FUNCTION F_RealToBitDword_1 : DWORD
VAR_INPUT
	rIn : REAL;
END_VAR
VAR
	pt : POINTER TO DWORD;
END_VAR

pt := ADR(rIn);
F_RealToBitDword := pt^;

END_FUNCTION

(* stored: Version 1.1.0.1, ProductVersion 3.1.4024.15
   POU F_RealToBitDword_1: Id {033f67c4-d697-408a-a5b9-465478a67f5e}, SpecialFunc None *)
